(* IEC 61131-3 sources: kns-pump-station/tests/POUs/Model/FB_StormGenerator_Test, 14 files *)

(* ---- FB_StormGenerator_Test.decl.st ---- *)
// Назначение: набор coUnit для FB_StormGenerator и F_Xorshift32 — ливни по seed: известные значения
//             xorshift32, ливни суток для seed по умолчанию, детерминизм и независимость от шага вызова,
//             трапеция, переход через полночь, снятие ливней, предел числа, нулевое состояние генератора.
//             Ожидаемые значения — эталон tools_project/plant_reference.py (сценарии xorshift.*, storms.*).
// Автор:      kr0nsch
// Версия:     0.1.0
// Документ:   docs/DESIGN.md, разделы 11.3, 14.1
FUNCTION_BLOCK FB_StormGenerator_Test EXTENDS coUnit.FB_TestSuite
VAR CONSTANT
    R_EPS_H : REAL := 1.0E-4;         // допуск начала ливня, ч (REAL против float64 эталона)
    R_EPS_M3H : REAL := 1.0E-3;       // допуск притока и пика, м³/ч
    UI_MAX_TOO_MANY : UINT := 10;     // больше SIM_STORMS_MAX
    UI_STEPS : UINT := 50;            // шагов часов в проверке независимости от шага
END_VAR

(* ---- ClearSuppressesRunningStorms.method.decl.st ---- *)
// Clear (xResetPlant) снимает идущий ливень и внеочередной ливень; ливни, которые начнутся позже
// (сутки 1, 4,80 ч), идут.
METHOD PRIVATE ClearSuppressesRunningStorms
VAR
    fbDut : FB_StormGenerator;  // проверяемый генератор
    stCfg : ST_SimCfg;          // параметры ливней по умолчанию
END_VAR

(* ---- CountLimitedToMax.method.decl.st ---- *)
// uiStormsPerDayMax = 10 ограничивается SIM_STORMS_MAX = 4 (эталон: по 4 ливня в сутки 0…2).
METHOD PRIVATE CountLimitedToMax
VAR
    fbDut : FB_StormGenerator;  // проверяемый генератор
    stCfg : ST_SimCfg;          // параметры ливней по умолчанию
END_VAR

(* ---- DefaultsSeedDayZeroStorms.method.decl.st ---- *)
// Параметры по умолчанию, сутки 0: два ливня — 2,7587 ч, 1 549 386 мс, 133,93 м³/ч и 4,5323 ч,
// 3 011 220 мс, 193,78 м³/ч; в 0 ч ливня нет.
METHOD PRIVATE DefaultsSeedDayZeroStorms
VAR
    fbDut : FB_StormGenerator;  // проверяемый генератор
    stCfg : ST_SimCfg;          // параметры ливней по умолчанию
END_VAR

(* ---- DifferentDaysDiffer.method.decl.st ---- *)
// Ливни разных суток и разных seed различаются (сутки 0 и 1; seed и seed + 1).
METHOD PRIVATE DifferentDaysDiffer
VAR
    fbDut : FB_StormGenerator;  // проверяемый генератор
    stCfg : ST_SimCfg;          // параметры ливней по умолчанию
    fbOther : FB_StormGenerator;
    rStartDay0 : REAL;          // начало первого ливня суток 0
END_VAR

(* ---- InflowDependsOnlyOnClock.method.decl.st ---- *)
// Приток зависит только от часов модели: 50 мелких шагов 4,5 → 5,0 ч и один вызов в 5,0 ч дают
// одинаковое значение (ливни одинаковы при любом ускорении); часы назад — значение как у нового
// генератора в том же моменте.
METHOD PRIVATE InflowDependsOnlyOnClock
VAR
    fbDut : FB_StormGenerator;  // проверяемый генератор
    stCfg : ST_SimCfg;          // параметры ливней по умолчанию
    fbOther : FB_StormGenerator;
    fbFresh : FB_StormGenerator;  // генератор, впервые вызванный в 4,6 ч
    uiK : UINT;
END_VAR

(* ---- InflowDependsOnlyOnClock.method.impl.st ---- *)
coUnit.TEST('StormGenerator_InflowDependsOnlyOnClock');

fbDut(lrClock_h := 4.5, udiSeed := stCfg.udiSeed, uiStormsPerDayMax := stCfg.uiStormsPerDayMax,
      rPeakMin_m3h := stCfg.rStormPeakMin_m3h, rPeakMax_m3h := stCfg.rStormPeakMax_m3h,
      tDurationMin := stCfg.tStormMin, tDurationMax := stCfg.tStormMax);
fbOther(lrClock_h := 5.0, udiSeed := stCfg.udiSeed, uiStormsPerDayMax := stCfg.uiStormsPerDayMax,
      rPeakMin_m3h := stCfg.rStormPeakMin_m3h, rPeakMax_m3h := stCfg.rStormPeakMax_m3h,
      tDurationMin := stCfg.tStormMin, tDurationMax := stCfg.tStormMax);
fbFresh(lrClock_h := 4.6, udiSeed := stCfg.udiSeed, uiStormsPerDayMax := stCfg.uiStormsPerDayMax,
      rPeakMin_m3h := stCfg.rStormPeakMin_m3h, rPeakMax_m3h := stCfg.rStormPeakMax_m3h,
      tDurationMin := stCfg.tStormMin, tDurationMax := stCfg.tStormMax);
FOR uiK := 1 TO UI_STEPS - 1 DO
    fbDut(lrClock_h := 4.5 + UINT_TO_LREAL(uiK) * 0.01);
END_FOR
fbDut(lrClock_h := 5.0);
AssertTrue(Condition := fbDut.rInflow_m3h > 0.0, Message := 'storm running at 5.0 h');
AssertEquals_REAL(Expected := fbOther.rInflow_m3h, Actual := fbDut.rInflow_m3h, Delta := 0.0,
                  Message := 'fine and coarse steps give same inflow');
fbDut(lrClock_h := 4.6);
AssertEquals_REAL(Expected := fbFresh.rInflow_m3h, Actual := fbDut.rInflow_m3h, Delta := 0.0,
                  Message := 'clock back: same inflow as fresh evaluation');

coUnit.TEST_FINISHED();

(* ---- SameSeedSameStorms.method.decl.st ---- *)
// Два генератора с одинаковым seed дают одинаковые ливни; сутки 1 совпадают с эталоном
// (4,8018 ч, 4 034 469 мс, 209,13 м³/ч и 0,3007 ч, 5 001 626 мс, 178,02 м³/ч).
METHOD PRIVATE SameSeedSameStorms
VAR
    fbDut : FB_StormGenerator;  // проверяемый генератор
    stCfg : ST_SimCfg;          // параметры ливней по умолчанию
    fbOther : FB_StormGenerator;  // второй генератор с тем же seed
    uiK : UINT;
END_VAR

(* ---- SameSeedSameStorms.method.impl.st ---- *)
coUnit.TEST('StormGenerator_SameSeedSameStorms');

fbDut(lrClock_h := 30.0, udiSeed := stCfg.udiSeed, uiStormsPerDayMax := stCfg.uiStormsPerDayMax,
      rPeakMin_m3h := stCfg.rStormPeakMin_m3h, rPeakMax_m3h := stCfg.rStormPeakMax_m3h,
      tDurationMin := stCfg.tStormMin, tDurationMax := stCfg.tStormMax);
fbOther(lrClock_h := 30.0, udiSeed := stCfg.udiSeed, uiStormsPerDayMax := stCfg.uiStormsPerDayMax,
      rPeakMin_m3h := stCfg.rStormPeakMin_m3h, rPeakMax_m3h := stCfg.rStormPeakMax_m3h,
      tDurationMin := stCfg.tStormMin, tDurationMax := stCfg.tStormMax);
AssertEquals_UDINT(Expected := 1, Actual := fbDut.udiDay, Message := 'day 1');
AssertEquals_UINT(Expected := fbDut.uiCount, Actual := fbOther.uiCount, Message := 'same count');
FOR uiK := 1 TO fbDut.uiCount DO
    AssertEquals_REAL(Expected := fbDut.astStorm[uiK].rStart_h, Actual := fbOther.astStorm[uiK].rStart_h, Delta := 0.0,
                      Message := 'same start');
    AssertEquals_TIME(Expected := fbDut.astStorm[uiK].tDuration, Actual := fbOther.astStorm[uiK].tDuration,
                      Message := 'same duration');
    AssertEquals_REAL(Expected := fbDut.astStorm[uiK].rPeak_m3h, Actual := fbOther.astStorm[uiK].rPeak_m3h,
                      Delta := 0.0,
                      Message := 'same peak');
END_FOR
// ref: storms.day1.*
AssertEquals_UINT(Expected := 2, Actual := fbDut.uiCount, Message := 'two storms on day 1');
AssertEquals_REAL(Expected := 4.801848, Actual := fbDut.astStorm[1].rStart_h, Delta := R_EPS_H,
                  Message := 'd1 s1 start');
AssertEquals_TIME(Expected := T#4034469MS, Actual := fbDut.astStorm[1].tDuration, Message := 'd1 s1 duration');
AssertEquals_REAL(Expected := 209.133103, Actual := fbDut.astStorm[1].rPeak_m3h, Delta := R_EPS_M3H,
                  Message := 'd1 s1 peak');
AssertEquals_REAL(Expected := 0.300672, Actual := fbDut.astStorm[2].rStart_h, Delta := R_EPS_H,
                  Message := 'd1 s2 start');
AssertEquals_TIME(Expected := T#5001626MS, Actual := fbDut.astStorm[2].tDuration, Message := 'd1 s2 duration');
AssertEquals_REAL(Expected := 178.015715, Actual := fbDut.astStorm[2].rPeak_m3h, Delta := R_EPS_M3H,
                  Message := 'd1 s2 peak');

coUnit.TEST_FINISHED();

(* ---- StormCrossingMidnightContinues.method.decl.st ---- *)
// Ливень суток 21 (23,8694 ч, 2 385 650 мс, 175,0 м³/ч) не закончился к полуночи: в 00:15 суток 22
// приток — его полка 175,0 м³/ч.
METHOD PRIVATE StormCrossingMidnightContinues
VAR
    fbDut : FB_StormGenerator;  // проверяемый генератор
    stCfg : ST_SimCfg;          // параметры ливней по умолчанию
    uiK : UINT;
    xFound : BOOL;              // ливень суток 21 найден
END_VAR

(* ---- StormCrossingMidnightContinues.method.impl.st ---- *)
coUnit.TEST('StormGenerator_StormCrossingMidnightContinues');

fbDut(lrClock_h := 527.0, udiSeed := stCfg.udiSeed, uiStormsPerDayMax := stCfg.uiStormsPerDayMax,
      rPeakMin_m3h := stCfg.rStormPeakMin_m3h, rPeakMax_m3h := stCfg.rStormPeakMax_m3h,
      tDurationMin := stCfg.tStormMin, tDurationMax := stCfg.tStormMax);
FOR uiK := 1 TO fbDut.uiCount DO
    IF ABS(fbDut.astStorm[uiK].rStart_h - 23.869357) < R_EPS_H THEN
        xFound := TRUE;
        AssertEquals_TIME(Expected := T#2385650MS, Actual := fbDut.astStorm[uiK].tDuration, Message := 'd21 duration');
    END_IF
END_FOR
// ref: storms.midnight_day21.*
AssertTrue(Condition := xFound, Message := 'day 21 storm at 23.8694 h');
fbDut(lrClock_h := 528.25);
AssertEquals_UDINT(Expected := 22, Actual := fbDut.udiDay, Message := 'day 22');
AssertTrue(Condition := fbDut.xActive, Message := 'storm continues after midnight');
AssertEquals_REAL(Expected := 174.999204, Actual := fbDut.rInflow_m3h, Delta := R_EPS_M3H,
                  Message := 'plateau after midnight');

coUnit.TEST_FINISHED();

(* ---- TrapezoidShape.method.decl.st ---- *)
// Внеочередной ливень (StartNow) 1 ч, пик 200 м³/ч: 4,5 мин — 100 (половина роста 15 %), 9 мин —
// 200, 30 мин — 200, 49,5 мин — 100 (половина спада 35 %), 60 мин — 0, ливень закончился.
METHOD PRIVATE TrapezoidShape
VAR
    fbDut : FB_StormGenerator;  // проверяемый генератор
    stCfg : ST_SimCfg;          // параметры ливней по умолчанию
END_VAR

(* ---- XorshiftKnownValues.method.decl.st ---- *)
// F_Xorshift32: из 1 — 270369 (Marsaglia, 2003); из seed по умолчанию 20261016 — 552152043, затем
// 3072158977 (эталон).
METHOD PRIVATE XorshiftKnownValues
VAR
    dwX : DWORD;                // состояние генератора
END_VAR

(* ---- ZeroSeedDoesNotStall.method.decl.st ---- *)
// seed 0 в сутки 0 даёт нулевое состояние xorshift — оно заменяется SIM_XS_ZERO_STATE; ливни
// детерминированы (эталон, до 4 в сутки: сутки 0 — 0, сутки 3 — 1, сутки 5 — 4).
METHOD PRIVATE ZeroSeedDoesNotStall
VAR
    fbDut : FB_StormGenerator;  // проверяемый генератор
    stCfg : ST_SimCfg;          // параметры ливней по умолчанию
END_VAR
